(* IEC 61131-3 sources: codesys-ai-industrial-robot-control/plc/src/Process/FB_PartTracker, 8 files *)

(* ---- CurrentX.st ---- *)
// Current belt-frame X of the part in slot uiIdx [mm].
METHOD CurrentX : LREAL
VAR_INPUT
    uiIdx : UINT;
END_VAR
VAR
    stR : ST_PartRecord;
END_VAR

stR := fbQueue.GetRecord(uiIdx);
CurrentX := stR.lrX + (lrBeltPos - stR.lrBeltPosAtCapture);

(* ---- Decide.st ---- *)
// Selects the bin, marks the record Decided and stores it.
METHOD PRIVATE Decide
VAR_INPUT
    uiIdx : UINT;
    stRecIn : ST_PartRecord;
END_VAR
VAR
    stOut : ST_PartRecord;
END_VAR

stOut := stRecIn;
stOut.eTargetBin := F_SelectBin(stOut, GVL_Params.rConfidenceThreshold, GVL_Params.aClassToBin);
stOut.eState := E_PartState.Decided;
IF stOut.xVisionValid AND stOut.rConfidence < GVL_Params.rConfidenceThreshold THEN
    RaiseEventAlarm(E_AlarmId.LowConfidence);
END_IF
fbQueue.PutRecord(uiIdx, stOut);

(* ---- FindPart.st ---- *)
// Slot index of the part with this id, or 0.
METHOD FindPart : UINT
VAR_INPUT
    udiPartId : UDINT;
END_VAR

FindPart := fbQueue.FindIndex(udiPartId);

(* ---- GetRecord.st ---- *)
METHOD GetRecord : ST_PartRecord
VAR_INPUT
    uiIdx : UINT;
END_VAR

GetRecord := fbQueue.GetRecord(uiIdx);

(* ---- NextPickable.st ---- *)
// The decided, identified part furthest downstream inside [lrMinX, lrMaxX] (belt frame), or 0.
METHOD NextPickable : UINT
VAR_INPUT
    lrMinX : LREAL;
    lrMaxX : LREAL;
END_VAR
VAR
    k : UINT;
    lrX : LREAL;
    lrBest : LREAL;
    stR : ST_PartRecord;
END_VAR

NextPickable := 0;
lrBest := lrMinX;
FOR k := 1 TO GVL_Config.MAX_PARTS DO
    stR := fbQueue.GetRecord(k);
    // a part vision did not see has no known class and height: it is not picked blind
    IF stR.eState = E_PartState.Decided AND stR.xVisionValid THEN
        lrX := CurrentX(k);
        IF lrX >= lrBest AND lrX <= lrMaxX THEN
            lrBest := lrX;
            NextPickable := k;
        END_IF
    END_IF
END_FOR

(* ---- RaiseAlarm.st ---- *)
METHOD PRIVATE RaiseAlarm
VAR_INPUT
    eId : E_AlarmId;
END_VAR

IF itfAlarms <> 0 THEN
    itfAlarms.Raise(eId);
END_IF

(* ---- RaiseEventAlarm.st ---- *)
METHOD PRIVATE RaiseEventAlarm
VAR_INPUT
    eId : E_AlarmId;
END_VAR

IF itfAlarms <> 0 THEN
    itfAlarms.RaiseEvent(eId);
END_IF

(* ---- SetState.st ---- *)
// Updates a part's state. Placed, Dropped and Missed parts are counted and their slot is freed;
// a missed part raises the PartMissed event.
METHOD SetState
VAR_INPUT
    uiIdx : UINT;
    eState : E_PartState;
END_VAR
VAR
    stR : ST_PartRecord;
END_VAR

stR := fbQueue.GetRecord(uiIdx);
IF stR.eState = E_PartState.Free THEN
    RETURN;
END_IF
CASE eState OF
    E_PartState.Placed:
        udiPlaced := udiPlaced + 1;
        fbQueue.Release(uiIdx);
    E_PartState.Dropped:
        udiDropped := udiDropped + 1;
        fbQueue.Release(uiIdx);
    E_PartState.Missed:
        udiMissed := udiMissed + 1;
        RaiseEventAlarm(E_AlarmId.PartMissed);
        fbQueue.Release(uiIdx);
ELSE
    stR.eState := eState;
    fbQueue.PutRecord(uiIdx, stR);
END_CASE
